(* IEC 61131-3 sources: llm-plc-st-eval/data/definitivo/gemini-3.1-pro-preview/A3/few_shot, 3 files *)

(* ---- ejec_1.st ---- *)
FUNCTION_BLOCK FB_Com
VAR_INPUT
    txReq : BOOL;   (* Peticion de transmision *)
    rxOk : BOOL;    (* Confirmacion de recepcion *)
    rxData : INT;   (* Dato recibido (eco) *)
END_VAR
VAR_OUTPUT
    txData : INT;   (* Dato a transmitir *)
    ocupado : BOOL; (* Intercambio en curso *)
    ok : BOOL;      (* Intercambio correcto *)
    error : BOOL;   (* Intercambio fallido tras 3 intentos *)
    nIntentos : INT;(* Numero de intento actual *)
END_VAR
VAR
    rTrigReq : R_TRIG; (* Detector de flanco para txReq *)
    rTrigRx : R_TRIG;  (* Detector de flanco para rxOk *)
    tTimeout : TON;    (* Temporizador de 500 ms *)
END_VAR

(* Deteccion de flancos *)
rTrigReq(CLK := txReq);
rTrigRx(CLK := rxOk);

(* Inicio de un nuevo intercambio si no hay uno en curso *)
IF rTrigReq.Q AND NOT ocupado THEN
    txData := 100;
    ocupado := TRUE;
    ok := FALSE;
    error := FALSE;
    nIntentos := 1;
    tTimeout(IN := FALSE, PT := T#500MS); (* Asegura el reinicio del temporizador *)
END_IF;

(* Control del intercambio en curso *)
IF ocupado THEN
    (* Actualiza el temporizador del intento actual *)
    tTimeout(IN := TRUE, PT := T#500MS);

    (* Evaluacion de la respuesta *)
    IF rTrigRx.Q AND (rxData = txData) THEN
        (* Intento correcto *)
        ok := TRUE;
        ocupado := FALSE;
        tTimeout(IN := FALSE, PT := T#500MS);

    ELSIF tTimeout.Q OR (rTrigRx.Q AND (rxData <> txData)) THEN
        (* Intento fallido por timeout o dato incorrecto *)
        IF nIntentos < 3 THEN
            (* Pasa al siguiente intento *)
            nIntentos := nIntentos + 1;
            tTimeout(IN := FALSE, PT := T#500MS); (* Reinicia el tiempo para el nuevo intento *)
        ELSE
            (* Fallaron los 3 intentos *)
            error := TRUE;
            ocupado := FALSE;
            tTimeout(IN := FALSE, PT := T#500MS);
        END_IF;
    END_IF;
END_IF;
END_FUNCTION_BLOCK

(* ---- ejec_2.st ---- *)
FUNCTION_BLOCK FB_Com
VAR_INPUT
    txReq : BOOL;  (* Peticion de transmision *)
    rxOk : BOOL;   (* Confirmacion de recepcion *)
    rxData : INT;  (* Datos recibidos (eco) *)
END_VAR
VAR_OUTPUT
    txData : INT;  (* Datos a transmitir *)
    ocupado : BOOL;(* Intercambio en curso *)
    ok : BOOL;     (* Intercambio correcto *)
    error : BOOL;  (* Intercambio fallido tras 3 intentos *)
    nIntentos : INT; (* Numero de intento actual *)
END_VAR
VAR
    flancoReq : R_TRIG; (* Detector de flanco para txReq *)
    flancoRx : R_TRIG;  (* Detector de flanco para rxOk *)
    temporizador : TON; (* Temporizador de 500 ms *)
    resetTemp : BOOL;   (* Señal para reiniciar el temporizador *)
END_VAR

(* Deteccion de flancos *)
flancoReq(CLK := txReq);
flancoRx(CLK := rxOk);

(* Inicio de un nuevo intercambio si no esta ocupado *)
IF flancoReq.Q AND NOT ocupado THEN
    ocupado := TRUE;
    ok := FALSE;
    error := FALSE;
    nIntentos := 1;
    txData := 100;
    resetTemp := TRUE;
ELSE
    resetTemp := FALSE;
END_IF;

(* Temporizador del intento en curso (se reinicia con resetTemp) *)
temporizador(IN := ocupado AND NOT resetTemp, PT := T#500MS);

(* Logica durante el intercambio *)
IF ocupado THEN
    (* Evaluacion de la respuesta *)
    IF flancoRx.Q THEN
        IF rxData = txData THEN
            (* Respuesta correcta (eco valido) *)
            ok := TRUE;
            ocupado := FALSE;
        ELSE
            (* Respuesta incorrecta: falla el intento *)
            IF nIntentos < 3 THEN
                nIntentos := nIntentos + 1;
                resetTemp := TRUE;
            ELSE
                error := TRUE;
                ocupado := FALSE;
            END_IF;
        END_IF;
    (* Evaluacion del timeout *)
    ELSIF temporizador.Q THEN
        IF nIntentos < 3 THEN
            nIntentos := nIntentos + 1;
            resetTemp := TRUE;
        ELSE
            error := TRUE;
            ocupado := FALSE;
        END_IF;
    END_IF;
END_IF;
END_FUNCTION_BLOCK

(* ---- ejec_3.st ---- *)
FUNCTION_BLOCK FB_Com
VAR_INPUT
    txReq : BOOL; (* Peticion de transmision *)
    rxOk : BOOL; (* Confirmacion de recepcion *)
    rxData : INT; (* Dato recibido (eco) *)
END_VAR
VAR_OUTPUT
    txData : INT; (* Dato a transmitir *)
    ocupado : BOOL; (* Intercambio en curso *)
    ok : BOOL; (* Intercambio finalizado con exito *)
    error : BOOL; (* Intercambio fallido tras 3 intentos *)
    nIntentos : INT; (* Numero de intento en curso *)
END_VAR
VAR
    reqTrig : R_TRIG; (* Flanco de subida de la peticion *)
    rxTrig : R_TRIG; (* Flanco de subida de la recepcion *)
    tTimeout : TON; (* Temporizador de plazo de espera *)
    resetTimer : BOOL; (* Pulso para reiniciar el temporizador *)
END_VAR

(* Deteccion de flancos *)
reqTrig(CLK := txReq);
rxTrig(CLK := rxOk);

(* Inicio de un nuevo intercambio (se ignora si ya esta ocupado) *)
IF reqTrig.Q AND NOT ocupado THEN
    txData := 100;
    ocupado := TRUE;
    ok := FALSE;
    error := FALSE;
    nIntentos := 1;
    resetTimer := TRUE;
END_IF;

(* Evaluacion del intento en curso *)
IF ocupado THEN
    IF rxTrig.Q AND (rxData = txData) THEN
        (* Confirmacion recibida correctamente *)
        ok := TRUE;
        ocupado := FALSE;
    ELSIF rxTrig.Q OR tTimeout.Q THEN
        (* Falla por dato incorrecto o por agotarse el tiempo (timeout) *)
        IF nIntentos < 3 THEN
            nIntentos := nIntentos + 1;
            resetTimer := TRUE; (* Reinicia el temporizador para el siguiente intento *)
        ELSE
            (* Se agotaron los 3 intentos *)
            error := TRUE;
            ocupado := FALSE;
        END_IF;
    END_IF;
END_IF;

(* Control del temporizador: se detiene si no esta ocupado o si se requiere reinicio *)
tTimeout(IN := ocupado AND NOT resetTimer, PT := T#500MS);
resetTimer := FALSE;

END_FUNCTION_BLOCK
